(* IEC 61131-3 sources: daoli-st-library/DL_Device, 362 files *)

(* ---- FB_DL_AnalogInputRedundancySel.st ---- *)
(*==============================================================================
 * 组件名称 (Component)  : FB_DL_AnalogInputRedundancySel
 * 所属子库 (Sublibrary) : DL_Device
 * 当前版本 (Version)    : 1.0.0
 * 兼容性   (Platform)   : CODESYS 3.5 / TwinCAT 3 / 汇川 InoProShop / 施耐德 Machine Expert
 *                         仅依赖 IEC 61131-3 标准库（ABS / MAX / MIN），零厂商方言
 * 功能描述 (Function)   : 双路模拟量冗余选择（无扰切换 + 偏差监控 + 坏值剔除）：
 *                         ① 两路均有效且 |A − B| ≤ fDevTol → 输出两路均值，选通码 3；
 *                         ② 两路均有效但偏差超限 → **按上一拍选定通道保持**（无扰切换），
 *                            置 bDevAlarm 与信息码，绝不两侧来回跳；
 *                         ③ 仅一路有效（另一路非有限 / 超量程）→ 剔除坏路、使用好路，
 *                            bChanAValid / bChanBValid 回执逐路披露；
 *                         ④ **双路皆坏 → eFault**：输出保持**上一有效值**，bValid=FALSE，
 *                            故障级码配对置 bError，恢复路径唯一：bReset 且至少一路恢复有效。
 * 接口     (Interface)  : 输入 8 项（使能 / 复位 / 两路原值 / 偏差容差 / 量程上下限），
 *                         输出 10 项（输出值 / 选通码 / 偏差告警 / 两路有效回执 /
 *                         状态回执 / 有效性与故障码）。
 * 边界     (Boundary)   : ① 量程判定用 [fRangeMin, fRangeMax] 闭区间，超界即该路无效
 *                            （不做单侧饱和，饱和会把坏值伪装成合法满量程）；
 *                         ② 偏差容差以 1E-9 为下限钳位，防零容差导致恒告警；
 *                         ③ 双路皆坏时输出保持 fLastValid（上一有效值），若从未有过
 *                            有效值则输出 0 哨兵并披露（bValid=FALSE）；
 *                         ④ 非有限双判：NaN 用 x <> x，Inf 用 |x − x| > EPS 双侧直比；
 *                         ⑤ 零全局耦合（无 GVL / VAR_EXTERNAL / %I / %Q）。
 * 码表     (Codes)      : 本件占用 16#0004_1020 ~ 16#0004_102F 区间，实际使用 5 个：
 *                         1020 信息级 容差/量程参数钳位；1021 信息级 仅单路有效已剔除坏路；
 *                         1022 信息级 双路偏差超限已保持上一通道；1023 故障级 双路皆坏；
 *                         1024 故障级 非法状态兜底。信息级码永不置 bError。
 * 分工声明 (Scope)      : 与 FB_DL_AnalogTransmitter 分工：那件做单路原始量→工程量的
 *                         标定与滤波；本件只做「两路冗余仲裁与坏值剔除」，不做标定。
 * 开源溯源 (Origin)     : 开源溯源：原创实现（无外部代码引入）
 * 红线自检 (Redline)    : R1 ✓ 零 GVL / VAR_EXTERNAL ｜ R2 ✓ 零 %I/%Q/%M
 *                         R3 ✓ 纯 IEC 61131-3 ｜ R4 ✓ 非有限双判 + 容差钳位 + 无除零
 *                         R5 ✓ 声明逐行同行双语注释 ｜ R6 ✓ 五态 ENUM + CASE + ELSE
 *                         R7 ✓ 无定时器/边沿实例（N/A），无跨周期定时依赖
 * 修订历史 (Revision)   : 2026-11-23  v1.0.0  R77 首版
 * 验收向量 (Acceptance) :
 *   V1 两路 A=10.0、B=10.4、fDevTol=1.0：fOut=10.2、iSelChan=3、bDevAlarm=FALSE、bValid=TRUE。
 *   V2 承接 V1，随后 A=10.0、B=15.0（偏差 5.0 > 1.0）：fOut 保持通道 A 的 10.0、
 *      iSelChan=1、bDevAlarm=TRUE、uErrorId=16#0004_1022、bError=FALSE（信息级）。
 *   V3 A=NaN、B=12.0：bChanAValid=FALSE、bChanBValid=TRUE、fOut=12.0、iSelChan=2、
 *      uErrorId=16#0004_1021、bError=FALSE。
 *   V4 A=NaN、B 超量程（B=200.0，量程上限 100.0）：双路皆坏 → eStateOut=eFault、
 *      fOut 保持上一有效值、bValid=FALSE、uErrorId=16#0004_1023、bError=TRUE。
 *   V5 承接 V4，bReset 单拍且 A 恢复为 10.0：eStateOut 回 eAvg/eHoldA，bError=FALSE。
 *============================================================================*)

(*-----------------------------------------------------------------------------
 * 调用示例 (Instance guide)：
 *   声明于调用方 FB 的 VAR 区：fbRed : FB_DL_AnalogInputRedundancySel;
 *   每周期无条件调用：fbRed(bEnable := TRUE, bReset := xReset,
 *                           fChanA := stAi.fCh1, fChanB := stAi.fCh2,
 *                           fDevTol := 0.5, fRangeMin := 0.0, fRangeMax := 100.0);
 *   取用出口：fPv := fbRed.fOut;  IF NOT fbRed.bValid THEN 保持工艺安全动作。
 *   注意：iSelChan 为「上一拍选定通道」的唯一载体，请勿在外部改写。
 *----------------------------------------------------------------------------*)

(*-----------------------------------------------------------------------------
 * 枚举: E_DL_ArsState（归属 DL_Device，与 FB_DL_AnalogInputRedundancySel 同文件）
 * 含义: 冗余选择状态机的离散状态。eAvg 为双路均值相，eHoldA / eHoldB 为单路保持相，
 *       eFault 为双路皆坏的故障相（输出保持上一有效值）。
 *----------------------------------------------------------------------------*)
TYPE E_DL_ArsState :
(
    eInit  := 0,    // 首扫态：输出直接取可用路，建立首个有效值 / First scan: output takes a valid channel to build the first valid value
    eAvg   := 10,   // 均值态：两路有效且偏差合格，输出均值 / Averaging state: both valid and deviation within tolerance
    eHoldA := 20,   // 保持 A 态：仅 A 有效或偏差超限且上一拍选 A / Hold channel A, valid alone or deviation exceeded with A previously selected
    eHoldB := 30,   // 保持 B 态：仅 B 有效或偏差超限且上一拍选 B / Hold channel B, valid alone or deviation exceeded with B previously selected
    eFault := 99    // 故障相：双路皆坏，输出保持上一有效值，bValid=FALSE / Fault: both channels bad, holds last valid value
);
END_TYPE

(*==============================================================================
 * 功能块: FB_DL_AnalogInputRedundancySel
 * 调用约定: 每周期无条件调用一次；无定时器/边沿实例（R7 N/A），全部判据单拍完成。
 * 无扰语义: 通道间切换只发生在「上一拍选定通道仍然有效」的前提下；一旦选定通道
 *           失效才切到另一路，切回条件为原通道恢复有效（而非偏差合格），避免抖动。
 *============================================================================*)
FUNCTION_BLOCK FB_DL_AnalogInputRedundancySel
VAR_INPUT
    bEnable    : BOOL := FALSE;         // 使能，FALSE 时输出冻结并置 bValid=FALSE / Enable, FALSE freezes the output and clears bValid
    bReset     : BOOL := FALSE;         // 复位（电平有效），解除双路皆坏锁存 / Reset (level), clears the both-bad latch
    fChanA     : REAL := 0.0;           // A 路原始采样值 [EU] / Raw sample of channel A [EU]
    fChanB     : REAL := 0.0;           // B 路原始采样值 [EU] / Raw sample of channel B [EU]
    fDevTol    : REAL := 0.5;           // 两路允许偏差容差 [EU] / Allowed deviation between the two channels [EU]
    fRangeMin  : REAL := 0.0;           // 量程下限（闭区间）[EU] / Range lower bound, closed interval [EU]
    fRangeMax  : REAL := 100.0;         // 量程上限（闭区间）[EU] / Range upper bound, closed interval [EU]
END_VAR
VAR_OUTPUT
    fOut       : REAL;                  // 仲裁输出值（双路皆坏时保持上一有效值）[EU] / Arbitrated output, holds last valid on both-bad
    iSelChan   : INT;                   // 选通码：0=无 1=A 2=B 3=均值 [-] / Selection code: 0=none 1=A 2=B 3=mean
    bDevAlarm  : BOOL;                  // 双路偏差超限告警（信息级，不置 bError）/ Deviation alarm, info level, keeps bError FALSE
    bChanAValid: BOOL;                  // A 路有效回执（有限且在量程内）/ Channel A validity feedback, finite and in range
    bChanBValid: BOOL;                  // B 路有效回执（有限且在量程内）/ Channel B validity feedback, finite and in range
    eStateOut  : E_DL_ArsState;         // 状态机当前状态回执 [-] / Current state feedback
    bValid     : BOOL;                  // 输出可信标志，故障相为 FALSE / Output trustworthy flag, FALSE in the fault state
    bError     : BOOL;                  // 故障级标志，与 uErrorId 严格联动 / Fault-level flag, strictly coupled with uErrorId
    uErrorId   : UDINT;                 // 错误码，0 = 无码 / Error code, 0 = no code
END_VAR
VAR
    eState     : E_DL_ArsState;         // 内部状态 [-] / Internal state
    fDev       : REAL;                  // 两路实时偏差绝对值 [EU] / Absolute deviation between the two channels [EU]
    fLastValid : REAL;                  // 上一有效输出值，故障相保持用 [EU] / Last valid output, held in the fault state
    bHaveLast  : BOOL;                  // 是否已建立过有效值 / A valid value has been established
    bBothValid : BOOL;                  // 两路均有效 / Both channels valid
    bOnlyA     : BOOL;                  // 仅 A 有效 / Only channel A valid
    bOnlyB     : BOOL;                  // 仅 B 有效 / Only channel B valid
    bNoneValid : BOOL;                  // 两路皆无效 / Neither channel valid
    bDevOk     : BOOL;                  // 偏差在容差内 / Deviation inside tolerance
    bChanANaN  : BOOL;                  // A 路自反判 NaN 命中 / Channel A NaN by self-comparison
    bChanAInf  : BOOL;                  // A 路差自减判 Inf 命中 / Channel A infinity by self-subtraction
    bChanBNaN  : BOOL;                  // B 路自反判 NaN 命中 / Channel B NaN by self-comparison
    bChanBInf  : BOOL;                  // B 路差自减判 Inf 命中 / Channel B infinity by self-subtraction
    bFaultLatch: BOOL;                  // 双路皆坏锁存位 / Both-bad latch
    bRangeBad  : BOOL;                  // 量程参数非法标志 / Range parameter invalid flag
    fDevTolEff : REAL;                  // 钳位后的偏差容差 [EU] / Clamped deviation tolerance [EU]
    fRangeLo   : REAL;                  // 生效量程下限 [EU] / Effective range lower bound [EU]
    fRangeHi   : REAL;                  // 生效量程上限 [EU] / Effective range upper bound [EU]
    uInfoCode  : UDINT;                 // 信息级码暂存 / Info-level code scratch
END_VAR
VAR CONSTANT
    DL_ARS_OK    : UDINT := 16#0000_0000;  // 无码哨兵 / No-code sentinel
    DL_ARS_TOL   : REAL := 1.0E-9;         // 容差硬下限，防零容差恒告警 [EU] / Tolerance floor preventing permanent alarm [EU]
    DL_ARS_EPS   : REAL := 1.0E-9;         // 浮点比较容差（统一口径）/ Unified floating point comparison tolerance
    DL_ARS_ZERO  : REAL := 0.0;            // 零基准哨兵 / Zero reference sentinel
    DL_ARS_HALF  : REAL := 0.5;            // 均值折半系数 / Averaging half factor
    DL_ARS_RANGE_DEF : REAL := 100.0;      // 量程非法时的兜底上限 [EU] / Fallback upper bound when the range is invalid [EU]
END_VAR

(*------------------------------------------------------------------------------
 * 段 0｜参数域闸（不中断扫描）：量程必须 fRangeMax > fRangeMin，容差 ≥ 1E-9
 *      Parameter domain gate: range must be increasing, tolerance floored
 *-----------------------------------------------------------------------------*)
uInfoCode  := DL_ARS_OK;                                    // 信息码预置无码 / Preset no info code
bRangeBad  := FALSE;                                        // 量程非法标志预置 / Preset range-invalid flag FALSE

fDevTolEff := MAX(fDevTol, DL_ARS_TOL);                     // 容差下限钳位 [EU] / Tolerance floor [EU]
fRangeLo   := fRangeMin;                                    // 生效量程下限 [EU] / Effective lower bound [EU]
IF fRangeMax > fRangeMin THEN
    fRangeHi := fRangeMax;                                  // 量程合法原值生效 [EU] / Legal upper bound applied [EU]
ELSE
    fRangeHi   := fRangeLo + DL_ARS_RANGE_DEF;              // 量程倒挂：改用兜底上限，拒绝零宽量程 / Inverted range, fallback width
    bRangeBad  := TRUE;                                     // 记录量程非法 / Record the invalid range
    uInfoCode  := 16#0004_1020;                             // 信息级：量程参数已钳位 / Info: range parameter clamped
END_IF

(*------------------------------------------------------------------------------
 * 段 1｜逐路有效性判定：非有限（NaN 自反 / Inf 差自减）与超量程（闭区间）双闸
 *      Per-channel validity: non-finite double test plus closed-interval range gate
 *-----------------------------------------------------------------------------*)
bChanANaN := (fChanA <> fChanA);                                                          // A 路自反判 NaN / Channel A NaN by self-comparison
bChanAInf := ABS(fChanA - fChanA) > DL_ARS_EPS;                                           // A 路差自减判 Inf（双侧直比）/ Channel A infinity by self-subtraction
bChanAValid := NOT (bChanANaN OR bChanAInf)
               AND (fChanA >= fRangeLo) AND (fChanA <= fRangeHi);                          // A 路有效回执 / Channel A validity

bChanBNaN := (fChanB <> fChanB);                                                          // B 路自反判 NaN / Channel B NaN by self-comparison
bChanBInf := ABS(fChanB - fChanB) > DL_ARS_EPS;                                           // B 路差自减判 Inf（双侧直比）/ Channel B infinity by self-subtraction
bChanBValid := NOT (bChanBNaN OR bChanBInf)
               AND (fChanB >= fRangeLo) AND (fChanB <= fRangeHi);                          // B 路有效回执 / Channel B validity

bBothValid := bChanAValid AND bChanBValid;                  // 两路均有效 / Both valid
bOnlyA     := bChanAValid AND (NOT bChanBValid);            // 仅 A 有效 / Only A valid
bOnlyB     := bChanBValid AND (NOT bChanAValid);            // 仅 B 有效 / Only B valid
bNoneValid := (NOT bChanAValid) AND (NOT bChanBValid);      // 两路皆无效 / Neither valid

(* 偏差只在两路都有效时才有意义；任一路坏时偏差保持上一拍值（不拿坏值重算）*)
(* The deviation is meaningful only when both channels are valid, otherwise it is held *)
IF bBothValid THEN
    fDev := ABS(fChanA - fChanB);                           // 两路偏差绝对值 [EU] / Absolute deviation [EU]
END_IF
bDevOk := bBothValid AND (fDev <= fDevTolEff);             // 偏差合格判据 [EU] / Deviation predicate [EU]

(*------------------------------------------------------------------------------
 * 段 2｜双路皆坏锁存：置位在 eFault 判断处，解除路径唯一：bReset 且至少一路有效
 *      Both-bad latch: cleared only by reset with at least one channel valid again
 *-----------------------------------------------------------------------------*)
IF bFaultLatch THEN
    IF bReset AND (bChanAValid OR bChanBValid) THEN
        bFaultLatch := FALSE;                               // 唯一解除路径：复位且至少一路恢复有效 / Sole clear path
    END_IF
ELSIF bNoneValid AND bEnable THEN
    bFaultLatch := TRUE;                                    // 双路皆坏：锁存 / Both channels bad, latch it
END_IF

(*------------------------------------------------------------------------------
 * 段 3｜主状态机（红线 R6）：ENUM + CASE + ELSE 兜底
 *      Main state machine with enum, case coverage and ELSE interception
 *      出口预置：本件所有分支都显式给 fOut / iSelChan / bValid，无隐式保持
 *-----------------------------------------------------------------------------*)
CASE eState OF

    eInit:
        (* 首扫：不做仲裁，直接取可用路建立首个有效值 *)
        (* First scan: no arbitration, take an available channel to build the first valid value *)
        bDevAlarm := FALSE;                                 // 告警复位 / Alarm reset
        IF bBothValid THEN
            fOut       := (fChanA + fChanB) * DL_ARS_HALF;  // 两路可用取均值 [EU] / Both usable, take the mean [EU]
            iSelChan   := 3;                                // 选通码 3 = 均值 / Selection code three, mean
            fLastValid := fOut;                             // 建立首个有效值 / Build the first valid value
            bHaveLast  := TRUE;                             // 有效值已建立 / Valid value established
            bValid     := TRUE;                             // 输出可信 / Output trustworthy
            eState     := eAvg;                             // 进均值相 / Enter the averaging state
        ELSIF bOnlyA THEN
            fOut       := fChanA;                           // 仅 A 可用 [EU] / Only A usable [EU]
            iSelChan   := 1;                                // 选通码 1 = A / Selection code one, A
            fLastValid := fOut;                             // 建立首个有效值 / Build the first valid value
            bHaveLast  := TRUE;                             // 有效值已建立 / Valid value established
            bValid     := TRUE;                             // 输出可信 / Output trustworthy
            eState     := eHoldA;                           // 进保持 A 相 / Enter hold A
        ELSIF bOnlyB THEN
            fOut       := fChanB;                           // 仅 B 可用 [EU] / Only B usable [EU]
            iSelChan   := 2;                                // 选通码 2 = B / Selection code two, B
            fLastValid := fOut;                             // 建立首个有效值 / Build the first valid value
            bHaveLast  := TRUE;                             // 有效值已建立 / Valid value established
            bValid     := TRUE;                             // 输出可信 / Output trustworthy
            eState     := eHoldB;                           // 进保持 B 相 / Enter hold B
        ELSIF bEnable THEN
            fOut      := fLastValid;                        // 双路皆坏：保持上一有效值（可能仍是 0 哨兵）/ Both bad, hold the last valid value
            iSelChan  := 0;                                 // 无选定通道 / No selected channel
            bValid    := FALSE;                             // 输出不可信 / Output untrustworthy
            bDevAlarm := FALSE;                             // 偏差判据不可得，不置告警 / Deviation unavailable, no alarm
            eState    := eFault;                            // 进故障相 / Enter the fault state
        ELSE
            fOut      := fLastValid;                        // 未使能：输出冻结 / Not enabled, output frozen
            iSelChan  := 0;                                 // 无选定通道 / No selected channel
            bValid    := FALSE;                             // 输出不可信 / Output untrustworthy
        END_IF

    eAvg:
        (* 均值相：两路仍有效且偏差合格才保持；偏差超限则保持上一拍选定通道 *)
        (* Averaging state: keep averaging while the deviation is fine, else hold the previous channel *)
        IF bNoneValid THEN
            fOut      := fLastValid;                        // 双路皆坏：保持上一有效值 / Both bad, hold the last valid value
            iSelChan  := 0;                                 // 无选定通道 / No selected channel
            bValid    := FALSE;                             // 输出不可信 / Output untrustworthy
            bDevAlarm := FALSE;                             // 偏差判据不可得 / Deviation unavailable
            eState    := eFault;                            // 进故障相 / Enter the fault state
        ELSIF bOnlyA THEN
            fOut       := fChanA;                           // 剔除坏路 B，用 A [EU] / Drop B, use A [EU]
            iSelChan   := 1;                                // 选通码 1 = A / Selection code one, A
            fLastValid := fOut;                             // 刷新上一有效值 / Refresh the last valid value
            bHaveLast  := TRUE;                             // 有效值已建立 / Valid value established
            bValid     := TRUE;                             // 输出可信 / Output trustworthy
            bDevAlarm  := FALSE;                            // 单路运行不属偏差告警 / Single-channel run is not a deviation alarm
            uInfoCode  := 16#0004_1021;                     // 信息级：仅单路有效已剔除坏路 / Info: single channel valid, bad one dropped
            eState     := eHoldA;                           // 进保持 A 相 / Enter hold A
        ELSIF bOnlyB THEN
            fOut       := fChanB;                           // 剔除坏路 A，用 B [EU] / Drop A, use B [EU]
            iSelChan   := 2;                                // 选通码 2 = B / Selection code two, B
            fLastValid := fOut;                             // 刷新上一有效值 / Refresh the last valid value
            bHaveLast  := TRUE;                             // 有效值已建立 / Valid value established
            bValid     := TRUE;                             // 输出可信 / Output trustworthy
            bDevAlarm  := FALSE;                            // 单路运行不属偏差告警 / Single-channel run is not a deviation alarm
            uInfoCode  := 16#0004_1021;                     // 信息级：仅单路有效已剔除坏路 / Info: single channel valid, bad one dropped
            eState     := eHoldB;                           // 进保持 B 相 / Enter hold B
        ELSIF bDevOk THEN
            fOut       := (fChanA + fChanB) * DL_ARS_HALF;  // 偏差合格：取均值 [EU] / Deviation fine, take the mean [EU]
            iSelChan   := 3;                                // 选通码 3 = 均值 / Selection code three, mean
            fLastValid := fOut;                             // 刷新上一有效值 / Refresh the last valid value
            bHaveLast  := TRUE;                             // 有效值已建立 / Valid value established
            bValid     := TRUE;                             // 输出可信 / Output trustworthy
            bDevAlarm  := FALSE;                            // 告警复位 / Alarm reset
        ELSE
            (* 偏差超限：无扰保持上一拍选定通道；均值相无历史通道时按 A 保持（口径写死）*)
            (* Deviation exceeded: hold the previous channel; from the mean state default to A *)
            fOut       := fChanA;                           // 保持 A 通道值（均值相缺历史时的固定口径）[EU] / Hold A, fixed policy from the mean state [EU]
            iSelChan   := 1;                                // 选通码 1 = A / Selection code one, A
            fLastValid := fOut;                             // 刷新上一有效值 / Refresh the last valid value
            bHaveLast  := TRUE;                             // 有效值已建立 / Valid value established
            bValid     := TRUE;                             // 输出可信 / Output trustworthy
            bDevAlarm  := TRUE;                             // 偏差超限告警置位 / Deviation alarm set
            uInfoCode  := 16#0004_1022;                     // 信息级：偏差超限已保持上一通道 / Info: deviation exceeded, previous channel held
            eState     := eHoldA;                           // 进保持 A 相 / Enter hold A
        END_IF

    eHoldA:
        (* 保持 A 相：A 仍有效即继续；A 失效则切 B；两路皆坏进故障相 *)
        (* Hold A: continue while A is valid, switch to B when A fails, fault when both bad *)
        IF bNoneValid THEN
            fOut      := fLastValid;                        // 双路皆坏：保持上一有效值 / Both bad, hold the last valid value
            iSelChan  := 0;                                 // 无选定通道 / No selected channel
            bValid    := FALSE;                             // 输出不可信 / Output untrustworthy
            bDevAlarm := FALSE;                             // 偏差判据不可得 / Deviation unavailable
            eState    := eFault;                            // 进故障相 / Enter the fault state
        ELSIF bChanAValid THEN
            fOut       := fChanA;                           // 保持 A 路 [EU] / Hold channel A [EU]
            iSelChan   := 1;                                // 选通码 1 = A / Selection code one, A
            fLastValid := fOut;                             // 刷新上一有效值 / Refresh the last valid value
            bHaveLast  := TRUE;                             // 有效值已建立 / Valid value established
            bValid     := TRUE;                             // 输出可信 / Output trustworthy
            IF bBothValid AND (NOT bDevOk) THEN
                bDevAlarm := TRUE;                          // 两路都在但偏差超限：维持告警 / Both valid but deviating, keep the alarm
                uInfoCode := 16#0004_1022;                  // 信息级：偏差超限保持通道 / Info: deviation exceeded, channel held
            ELSE
                bDevAlarm := FALSE;                         // 偏差回落清除告警 / Alarm cleared when the deviation settles
            END_IF
        ELSE
            fOut       := fChanB;                           // A 失效切 B（B 此时必然有效）[EU] / A failed, switch to B, which must be valid [EU]
            iSelChan   := 2;                                // 选通码 2 = B / Selection code two, B
            fLastValid := fOut;                             // 刷新上一有效值 / Refresh the last valid value
            bHaveLast  := TRUE;                             // 有效值已建立 / Valid value established
            bValid     := TRUE;                             // 输出可信 / Output trustworthy
            bDevAlarm  := FALSE;                            // 单路运行不属偏差告警 / Single-channel run is not a deviation alarm
            uInfoCode  := 16#0004_1021;                     // 信息级：仅单路有效已剔除坏路 / Info: single channel valid, bad one dropped
            eState     := eHoldB;                           // 进保持 B 相 / Enter hold B
        END_IF

    eHoldB:
        (* 保持 B 相：B 仍有效即继续；B 失效则切 A；两路皆坏进故障相 *)
        (* Hold B: continue while B is valid, switch to A when B fails, fault when both bad *)
        IF bNoneValid THEN
            fOut      := fLastValid;                        // 双路皆坏：保持上一有效值 / Both bad, hold the last valid value
            iSelChan  := 0;                                 // 无选定通道 / No selected channel
            bValid    := FALSE;                             // 输出不可信 / Output untrustworthy
            bDevAlarm := FALSE;                             // 偏差判据不可得 / Deviation unavailable
            eState    := eFault;                            // 进故障相 / Enter the fault state
        ELSIF bChanBValid THEN
            fOut       := fChanB;                           // 保持 B 路 [EU] / Hold channel B [EU]
            iSelChan   := 2;                                // 选通码 2 = B / Selection code two, B
            fLastValid := fOut;                             // 刷新上一有效值 / Refresh the last valid value
            bHaveLast  := TRUE;                             // 有效值已建立 / Valid value established
            bValid     := TRUE;                             // 输出可信 / Output trustworthy
            IF bBothValid AND (NOT bDevOk) THEN
                bDevAlarm := TRUE;                          // 两路都在但偏差超限：维持告警 / Both valid but deviating, keep the alarm
                uInfoCode := 16#0004_1022;                  // 信息级：偏差超限保持通道 / Info: deviation exceeded, channel held
            ELSE
                bDevAlarm := FALSE;                         // 偏差回落清除告警 / Alarm cleared when the deviation settles
            END_IF
        ELSE
            fOut       := fChanA;                           // B 失效切 A（A 此时必然有效）[EU] / B failed, switch to A, which must be valid [EU]
            iSelChan   := 1;                                // 选通码 1 = A / Selection code one, A
            fLastValid := fOut;                             // 刷新上一有效值 / Refresh the last valid value
            bHaveLast  := TRUE;                             // 有效值已建立 / Valid value established
            bValid     := TRUE;                             // 输出可信 / Output trustworthy
            bDevAlarm  := FALSE;                            // 单路运行不属偏差告警 / Single-channel run is not a deviation alarm
            uInfoCode  := 16#0004_1021;                     // 信息级：仅单路有效已剔除坏路 / Info: single channel valid, bad one dropped
            eState     := eHoldA;                           // 进保持 A 相 / Enter hold A
        END_IF

    eFault:
        (* 故障相：输出保持上一有效值，bValid=FALSE；恢复路径唯一：bReset 且至少一路有效 *)
        (* Fault: hold the last valid value, recover only via reset with one valid channel *)
        fOut      := fLastValid;                            // 保持上一有效值（从未有过则为 0 哨兵）/ Hold the last valid value
        iSelChan  := 0;                                     // 无选定通道 / No selected channel
        bValid    := FALSE;                                 // 输出不可信 / Output untrustworthy
        bDevAlarm := FALSE;                                 // 偏差判据不可得，不置告警 / Deviation unavailable, no alarm
        IF (NOT bEnable) THEN
            eState := eInit;                                // 失能回首扫态 / Disable returns to init
        ELSIF (NOT bFaultLatch) AND bChanAValid THEN
            eState := eHoldA;                               // 复位后 A 恢复有效 / A recovered after reset
        ELSIF (NOT bFaultLatch) AND bChanBValid THEN
            eState := eHoldB;                               // 复位后 B 恢复有效 / B recovered after reset
        END_IF

    ELSE
        (* 非法状态拦截：任何未定义枚举值一律进故障相并置兜底码 *)
        (* Illegal state interception: undefined enum values go to fault with a fallback code *)
        eState    := eFault;                                // 强制回故障相 / Force back to the fault state
        fOut      := fLastValid;                            // 输出保持上一有效值 / Output holds the last valid value
        iSelChan  := 0;                                     // 无选定通道 / No selected channel
        bValid    := FALSE;                                 // 输出不可信 / Output untrustworthy
        bDevAlarm := FALSE;                                 // 不置偏差告警 / No deviation alarm
        uInfoCode := 16#0004_1024;                          // 故障级：非法状态兜底 / Fault: illegal state fallback

END_CASE

(*------------------------------------------------------------------------------
 * 段 4｜无扰冻结：未使能时输出冻结在上一有效值（不跟随输入）
 *      Bumpless freeze: while disabled the output stays on the last valid value
 *-----------------------------------------------------------------------------*)
IF NOT bEnable THEN
    IF bHaveLast THEN
        fOut := fLastValid;                                 // 冻结在上一有效值 / Freeze on the last valid value
    ELSE
        fOut := DL_ARS_ZERO;                                // 从未有过有效值：输出 0 哨兵 / Never valid, emit the zero sentinel
    END_IF
    bValid    := FALSE;                                     // 冻结相输出不可信 / Frozen output is not trustworthy
    bDevAlarm := FALSE;                                     // 冻结相不产生告警 / No alarm while frozen
END_IF

(*------------------------------------------------------------------------------
 * 段 5｜故障码统一出口（故障级锁存回放，信息级不置 bError）
 *      Unified code outlet: fault codes replayed latched, info codes never raise bError
 *-----------------------------------------------------------------------------*)
IF bFaultLatch THEN
    uErrorId := 16#0004_1023;                               // 故障级：双路皆坏 / Fault: both channels bad
    bError   := TRUE;                                       // 故障级码配对置位 / Paired fault flag set
ELSIF uInfoCode = 16#0004_1024 THEN
    uErrorId := 16#0004_1024;                               // 故障级：非法状态兜底 / Fault: illegal state fallback
    bError   := TRUE;                                       // 故障级码配对置位 / Paired fault flag set
ELSE
    uErrorId := uInfoCode;                                  // 信息级码或 0 / Info code or zero
    bError   := FALSE;                                      // 信息级不置故障标志 / Info level never raises the fault flag
END_IF

eStateOut := eState;                                        // 状态回执单一出口 / State feedback through a single outlet
END_FUNCTION_BLOCK

(* ---- FB_DL_AnalogSignalHealth.st ---- *)
// ==============================================================================
// 组件名 Component  : FB_DL_AnalogSignalHealth
// 分类   Category   : DL_Device
// 前缀   Naming     : FB_DL_ ｜ b/f/e/t/u 类型前缀制（R265）
// 版本   Version    : 1.0.0
// 复杂度 Complexity  : 中
// 功能   Purpose    : 4-20mA 模拟量信号健康诊断：断线（< 3.6 mA）、超上限
//                      （> fSatHigh）、低限（fSatLow ≤ 值 < 3.6 之外的
//                      低带口径见边界三）、卡滞（变化率绝对值持续
//                      <= fStuckBand 超 tStuck）；报警锁存至 bReset 上升沿，
//                      沿脉冲单拍。供变送器回路质量监视与预测性维护。
// 开源溯源 Origin    : 西门子 LGF 分类语义借鉴，clean-room 重写（LGF
//                      Process Diagnostics「模拟量断线 / 饱和监视」分类学
//                      口径借鉴，只借骨不抄肉，判据与实现零代码复制）
// 许可证 License    : MIT
// 参考   Reference  : IEC 61131-3:2013 §6.6 TON / R_TRIG 语义；NAMUR
//                      NE43 信号电平分级公开条款（借 3.6/4/20/20.5 mA
//                      分级语义，不抄文）
// 平台   Platform   : 纯 IEC 61131-3（TON / R_TRIG / LREAL 比较），三平台通用
// 依赖   Depends    : 仅 Standard.library（TON / R_TRIG 属标准件）
// 分工声明 Split     : FB_DL_SignalStuckWatch（通用卡滞监视）/ FB_DL_Analog
//                      Transmitter（模拟量变换）与本件互引；本件为 4-20mA
//                      回路专属健康分级（NE43 口径 + 回路卡滞三合一），
//                      通用信号冻结监视归 SignalStuckWatch（R216）。
// 归属 Ownership     : E_DL_AshHealth 属主为本文件（全库唯一定义，R264）；
//                      引用件只引用不重声明。
// ------------------------------------------------------------------
// 边界 Boundary     :
//   一 TON 无条件刷新（R7）：tonStuck 于段 0 顶层调用，IN 串「有变化即
//      重置」口径——IN := 变化率绝对值 <= fStuckBand（有变化时 IN 为
//      FALSE 计时自清，卡滞即「无变化持续超窗」）；首拍 / 复位后
//      _bPrevValid = FALSE 不计时（防假前值参与变化率）；
//   二 判据分级（R190 归因唯一，独立码位）：fMa 非有限 → eInvalid
//      （bValid = FALSE 通道，无码位）；fMa < 3.6 → eWireBreak（断线）；
//      fMa >= 3.6 且 fMa < fSatLow → eSatLow（低限）；fMa > fSatHigh →
//      eSatHigh（超上限）；其余正常带内 tonStuck.Q → eStuck（卡滞）；
//      以上皆否 → eOk；
//   三 低限口径声明：3.6 mA 硬断线阈值与 fSatLow 组态阈值分离——
//      fSatLow 默认 3.6（与硬阈值重合），调用方可上调 fSatLow 收紧
//      低带；fSatLow 下调低于 3.6 时低限带被硬阈值吸收（合法组态）；
//   四 报警锁存：_bAlarmLatch 置位后保持至 bReset 上升沿（锁存解除式
//      可达自证：输入引脚恒可达，R152）；首报码 _uErrLatch 锁存回放
//      （FB33-1：不在故障态按当下输入重新推断）；bAlarmEdge 单拍
//      （新报警沿，已锁存期不再发）；
//   五 组态守卫（防御性补码，R272 逐项点名）：fSatLow >= fSatHigh、
//      fSatLow / fSatHigh / fStuckBand 非有限、fStuckBand < 0、
//      tStuck <= 0 任一成立 → eHealth = eInvalid、bValid = FALSE、
//      报警锁存（故障级 0735）；
//   六 卡滞窗与报警锁存互锁：_bAlarmLatch 期间 tonStuck.IN 强制 FALSE
//      （复位沿同拍不重锁，FB50-1），复位后 _bPrevValid 清零重练；
//   七 失能（bEn = FALSE）语义写死（R303 离相清零）：eHealth 回 eOk、
//      报警锁存 / 码锁存清零、bValid = FALSE（失能不是故障）；
//   八 无除法；无全局、无外部变量、无物理地址；无状态机 CASE
//      （IF 判据链，末位 ELSE 兜底为 eOk）。
// 错误码 Codes      :
//   16#0003_0201【信息级】断线（fMa < 3.6 mA，NE43 口径）→ eWireBreak
//   16#0003_0202【信息级】超上限（fMa > fSatHigh）→ eSatHigh
//   16#0003_0203【信息级】低限（3.6 ≤ fMa < fSatLow）→ eSatLow
//   16#0003_0204【信息级】卡滞（变化率 <= fStuckBand 持续 tStuck）→ eStuck
//   16#0003_0735【故障级】组态非法（fSatLow >= fSatHigh / 参数非有限 /
//                fStuckBand < 0 / tStuck <= 0）→ eInvalid + bValid = FALSE
//   注：0201~0204 段位按本轮任务定稿启用（信息级，经 eErr / bAlarm
//   通道表达）；fMa 非有限走 eInvalid 无码位（bValid = FALSE 通道）。
//   0201~0204 四码分立依据（R90）：处置人不同（断线查接线、超限查
//   量程组态、低限查供电、卡滞查管路 / 变送器膜片），场景互斥可还原。
// 验收 Acceptance   :
//   算法已证（脚本）：未跑 ｜ 编译器已证（三平台）：未跑
//   V1 fMa = 3.0 → eWireBreak + 码 0201 + bAlarm 锁存
//   V2 fMa = 21.0 → eSatHigh + 码 0202；fMa = 3.7（fSatLow = 4.0）→ eSatLow
//   V3 fMa 恒 12.000 ± 0.01 超 10s → eStuck + 码 0204
//   V4 fMa 恒定但 < 3.6 → 断线优先（卡滞窗被门控不计时）
//   V5 fMa = NaN → eInvalid + bValid = FALSE（无码位）
//   V6 bReset 上升沿 → 锁存清零、卡滞计时重练（_bPrevValid 清零）
//   V7 bEn = FALSE → 全出口清零回 eOk（R303）
//   V8 fSatLow = 25（>= fSatHigh）→ 0735 + eInvalid
// 修订记录 Revision  :
//   2026-11-22  v1.0.0  R65 首版（批 3 · 序号 9，LGF Process Diagnostics 补口）
// ==============================================================================
TYPE E_DL_AshHealth :
(
    eOk        := 0,  // 健康带内 / ok, the signal in the healthy band
    eWireBreak := 10, // 断线：fMa < 3.6 mA（NE43 口径）/ the wire break under the hard threshold
    eSatHigh   := 20, // 超上限：fMa > fSatHigh / the saturation above the configured high
    eSatLow    := 30, // 低限：3.6 <= fMa < fSatLow / the low limit under the configured low
    eStuck     := 40, // 卡滞：变化率持续不超带超窗 / the stuck value through the window
    eInvalid   := 50  // 无效：输入非有限或组态非法 / invalid, a non finite input or configuration
);
END_TYPE

FUNCTION_BLOCK FB_DL_AnalogSignalHealth
VAR_INPUT
    fMa        : LREAL;         // 实测电流 [mA]（4-20mA 回路）/ the measured current in milliamps
    bEn        : BOOL := TRUE;  // 使能 [-]，FALSE 时出口清零回 eOk（R303）/ the enable
    fSatLow    : LREAL := 3.6;  // 低限阈值 [mA]，须 < fSatHigh / the low limit threshold
    fSatHigh   : LREAL := 20.5; // 超上限阈值 [mA]，NE43 口径默认 20.5 / the saturation high threshold
    fStuckBand : LREAL := 0.05; // 卡滞变化带 [mA]，变化率绝对值 <= 此值视为无变化 / the stuck band of the rate
    tStuck     : TIME := T#10S; // 卡滞判定窗 [毫秒]，须 > 0 / the stuck window, above zero
    bReset     : BOOL := FALSE; // 报警复位电平，上升沿清锁存（边界四解除式）/ the reset level, its rising edge releases the latch
END_VAR
VAR_OUTPUT
    eHealth    : E_DL_AshHealth := E_DL_AshHealth.eOk; // 健康状态出口 [状态] / the health outlet
    bAlarm     : BOOL := FALSE; // 报警锁存 [-]，任一非 eOk 状态置位至复位 / the latched alarm
    bAlarmEdge : BOOL := FALSE; // 新报警沿脉冲 [-]，单拍有效 / the new alarm edge pulse, single scan
    bValid     : BOOL := FALSE; // 判据可用 [-]，输入非有限或组态非法为 FALSE / the criteria usable flag
    eErr       : UDINT := 16#0000_0000; // 错误码，0 = 正常（首报码锁存回放）/ the error code, zero is ok
END_VAR
VAR
    _fPrevMa     : LREAL := 0.0;  // 前拍 mA 快照 [mA]（卡滞变化率基准）/ the previous scan snapshot of fMa
    _bPrevValid  : BOOL := FALSE; // 前值有效标志 [-]（首拍 / 复位后不参与变化率）/ the previous value valid flag
    _bAlarmLatch : BOOL := FALSE; // 报警锁存副本 [-]（仅复位沿清除）/ the alarm latch copy
    _uErrLatch   : UDINT := 16#0000_0000; // 首报码锁存 [码]（复位沿清除，FB33-1）/ the latched first report code
    _bAlarmNew   : BOOL := FALSE; // 本拍新报警标志 [-]（沿脉冲源，单拍）/ the new alarm flag of this scan
    _eHealthInt  : E_DL_AshHealth := E_DL_AshHealth.eOk; // 健康状态内部判定 [状态] / the internal health verdict
    _uCodeNow    : UDINT := 16#0000_0000; // 本拍判据码 [码] / the verdict code of this scan
    _bMaBad      : BOOL;          // fMa 非有限标志（逐拍重算）/ the input fault flag
    _bCfgBad     : BOOL;          // 组态非法标志（逐拍重算）/ the configuration fault flag
    _bInBand     : BOOL;          // 处于正常工作带 [-]（卡滞计时前提）/ the in band flag, the stuck timer premise
    _bDeltaSmall : BOOL;          // 变化率不超带 [-]（卡滞计时条件）/ the small rate flag
    rtReset      : R_TRIG;        // 复位沿实例，段 0 无条件刷新（R7）/ the reset edge instance refreshed unconditionally
    tonStuck     : TON;           // 卡滞窗定时器，段 0 无条件刷新 / the stuck window timer refreshed unconditionally
END_VAR
VAR CONSTANT
    DL_ASH_WIRE  : LREAL := 3.6;            // 硬断线阈值 [mA]（NE43 口径）/ the hard wire break threshold
    DL_ASH_FMAX  : LREAL := 1.0E30;         // 非有限筛查幅值上限 [mA] / the finiteness screening cap
    DL_ASH_TIME0 : TIME := T#0S;            // 时间零常量 [毫秒] / the time zero constant
    DL_ASH_ZEROU : UDINT := 16#0000_0000;   // 码零常量 / the code zero constant
    DL_ASH_E_WIRE  : UDINT := 16#0003_0201; // 信息级：断线 / the wire break code
    DL_ASH_E_SATHI : UDINT := 16#0003_0202; // 信息级：超上限 / the saturation high code
    DL_ASH_E_SATLO : UDINT := 16#0003_0203; // 信息级：低限 / the low limit code
    DL_ASH_E_STUCK : UDINT := 16#0003_0204; // 信息级：卡滞 / the stuck code
    DL_ASH_E_CFG   : UDINT := 16#0003_0735; // 故障级：组态非法 / the configuration fault code
END_VAR

// 段 0｜定时器与沿实例无条件周期刷新（禁入分支，R7）/ segment 0, the unconditional refresh
rtReset(CLK := bReset);          // 复位沿 / the reset edge
_bMaBad := (fMa <> fMa) OR ((fMa - fMa) <> 0.0) OR (ABS(fMa) > DL_ASH_FMAX); // 输入非有限（NaN 自反判 + Inf 差值自反判 + 幅值上界，R272）/ the input non finite
_bCfgBad := (fSatLow >= fSatHigh)                                        // 低限不低于上限 / the low limit above the high
         OR (fSatLow <> fSatLow) OR ((fSatLow - fSatLow) <> 0.0) OR (ABS(fSatLow) > DL_ASH_FMAX)     // fSatLow 非有限 / fSatLow non finite
         OR (fSatHigh <> fSatHigh) OR ((fSatHigh - fSatHigh) <> 0.0) OR (ABS(fSatHigh) > DL_ASH_FMAX) // fSatHigh 非有限 / fSatHigh non finite
         OR (fStuckBand < 0.0)                                           // 变化带为负 / a negative band
         OR (fStuckBand <> fStuckBand) OR ((fStuckBand - fStuckBand) <> 0.0) OR (ABS(fStuckBand) > DL_ASH_FMAX) // fStuckBand 非有限 / fStuckBand non finite
         OR (tStuck <= DL_ASH_TIME0);                                    // 卡滞窗非正 / a non positive window
_bInBand := (NOT _bMaBad) AND (NOT _bCfgBad) AND (fMa >= DL_ASH_WIRE) AND (fMa >= fSatLow) AND (fMa <= fSatHigh); // 正常工作带（卡滞计时前提，边界二）/ the healthy band, the stuck timer premise
_bDeltaSmall := _bPrevValid AND (ABS(fMa - _fPrevMa) <= fStuckBand); // 变化率不超带（有变化时为 FALSE 计时自清，边界一）/ the rate within the band
tonStuck(IN := bEn AND _bInBand AND (NOT _bAlarmLatch) AND _bDeltaSmall, PT := tStuck); // 卡滞窗计时（串使能 / 带 / 锁存门控，FB50-1；锁存期 IN 强制 FALSE 防复位同拍重锁，边界六）/ the stuck window with the full gating

// 段 1｜单拍量预清零 + 复位沿作用域（R256 / R311）/ segment 1, the preset and the reset edge scope
bAlarmEdge := FALSE;             // 沿脉冲预清零（单拍信息位）/ preset the edge pulse false
IF rtReset.Q THEN                // 复位沿（作用域声明：清双锁存 + 重练卡滞计时，R311）/ the reset edge with the declared scope
    _bAlarmLatch := FALSE;       // 清报警锁存（唯一解除路径，边界四自证可达）/ clear the alarm latch
    _uErrLatch := DL_ASH_ZEROU;  // 清首报码锁存 / clear the latched code
    _bPrevValid := FALSE;        // 前值失效（卡滞计时重练，防旧基线误判）/ invalidate the previous value
    _fPrevMa := 0.0;             // 前值显式清零 [mA] / clear the previous value explicitly
END_IF

// 段 2｜失能分支：出口清零回 eOk，不 faults（R303 离相清零声明行）/ segment 2, the disabled branch
IF NOT bEn THEN                  // 失能 / disabled
    _eHealthInt := E_DL_AshHealth.eOk; // 强制健康态 / force the healthy state
    _bAlarmLatch := FALSE;       // 清报警锁存（使能断开 ≠ 信号故障）/ clear the alarm latch
    _uErrLatch := DL_ASH_ZEROU;  // 清码锁存 / clear the latched code
    _bPrevValid := FALSE;        // 前值失效（重新使能后重练）/ invalidate the previous value
    eHealth := _eHealthInt;      // 状态出口 / the health outlet
    bAlarm := FALSE;             // 报警位复位 / the alarm bit resets
    bAlarmEdge := FALSE;         // 沿脉冲复位 / the edge pulse resets
    bValid := FALSE;             // 失能即不可用 / not usable while disabled
    eErr := DL_ASH_ZEROU;        // 失能不发码 / no code while disabled
    RETURN;                      // 早退 / early return
END_IF

// 段 3｜判据分级链（边界二 / 五：R190 归因唯一，末位 ELSE 兜底 eOk）/ segment 3, the verdict chain
IF _bCfgBad THEN                 // 组态非法优先（故障级 0735）/ the configuration fault first
    _eHealthInt := E_DL_AshHealth.eInvalid; // 无效态 / the invalid state
    _uCodeNow := DL_ASH_E_CFG;   // 故障级码 / the fault code
ELSIF _bMaBad THEN               // 输入非有限 / a non finite input
    _eHealthInt := E_DL_AshHealth.eInvalid; // 无效态 / the invalid state
    _uCodeNow := DL_ASH_ZEROU;   // 无码位（bValid = FALSE 通道表达，边界二）/ no code, the validity channel speaks
ELSIF fMa < DL_ASH_WIRE THEN     // 硬断线阈值之下（NE43 口径）/ under the hard wire break threshold
    _eHealthInt := E_DL_AshHealth.eWireBreak; // 断线态 / the wire break state
    _uCodeNow := DL_ASH_E_WIRE;  // 信息级 0201 / the wire break code
ELSIF fMa < fSatLow THEN         // 低限带（fMa >= 3.6 已由上分支证明）/ the low limit band
    _eHealthInt := E_DL_AshHealth.eSatLow;   // 低限态 / the low limit state
    _uCodeNow := DL_ASH_E_SATLO; // 信息级 0203 / the low limit code
ELSIF fMa > fSatHigh THEN        // 超上限 / over the high threshold
    _eHealthInt := E_DL_AshHealth.eSatHigh;  // 超上限态 / the saturation state
    _uCodeNow := DL_ASH_E_SATHI; // 信息级 0202 / the saturation code
ELSIF tonStuck.Q THEN            // 卡滞超窗（正常带内才有资格判，边界二 / 六）/ stuck through the window
    _eHealthInt := E_DL_AshHealth.eStuck;    // 卡滞态 / the stuck state
    _uCodeNow := DL_ASH_E_STUCK; // 信息级 0204 / the stuck code
ELSE                             // 兜底：健康 / the fallback, healthy
    _eHealthInt := E_DL_AshHealth.eOk;       // 健康态 / the healthy state
    _uCodeNow := DL_ASH_ZEROU;   // 无码 / no code
END_IF

// 段 4｜报警锁存与首报码（边界四：锁存回放，FB33-1）/ segment 4, the alarm latch and the first report code
_bAlarmNew := FALSE;             // 新报警标志预清零 / preset the new alarm flag false
IF _eHealthInt <> E_DL_AshHealth.eOk THEN // 判据非健康 / the verdict not healthy
    IF NOT _bAlarmLatch THEN     // 首次报警 / a first alarm
        _bAlarmNew := TRUE;      // 置新报警标志（沿脉冲源，单拍）/ raise the new alarm flag
        _uErrLatch := _uCodeNow; // 首报码锁存（此后回放，不按当下输入重推断）/ latch the first code for the replay
    END_IF
    _bAlarmLatch := TRUE;        // 报警锁存至复位沿 / latch the alarm to the reset edge
END_IF

// 段 5｜统一出口（名实双出口同源，R191）/ segment 5, the unified outlet
eHealth := _eHealthInt;          // 状态出口 / the health outlet
bAlarm := _bAlarmLatch;          // 报警位与锁存同源 / the alarm bit from the latch
bAlarmEdge := _bAlarmNew;        // 沿脉冲单拍（已锁存期不再发）/ the single scan edge pulse
bValid := (NOT _bMaBad) AND (NOT _bCfgBad); // 判据可用（无输入 / 组态故障）/ usable without faults
IF _bAlarmLatch THEN             // 报警锁存回放优先 / the latched code replays first
    eErr := _uErrLatch;          // 首报码回放 / replay the latched code
ELSE                             // 无报警 / no alarm
    eErr := DL_ASH_ZEROU;        // 正常 / ok
END_IF

// 段 6｜前拍快照更新（边界一：仅有限值更新，非有限保旧值）/ segment 6, the previous value update
IF NOT _bMaBad THEN              // 输入有限才更新基准 / update the baseline only on a finite input
    _fPrevMa := fMa;             // 前拍快照刷新 [mA] / refresh the snapshot
    _bPrevValid := TRUE;         // 前值有效 / the previous value valid
END_IF
END_FUNCTION_BLOCK

(* ---- FB_DL_AxiolineDiagLatch.st ---- *)
(*==============================================================================
 * 组件名称 (Component)  : FB_DL_AxiolineDiagLatch
 * 所属子库 (Sublibrary) : DL_Device
 * 当前版本 (Version)    : 1.0.1
 * 组件分类 (Category)   : 功能块（FUNCTION_BLOCK）· 设备诊断 · 总线位域解析
 * 兼容性   (Platform)   : CODESYS 3.5 / TwinCAT 3 / 汇川 InoProShop / Schneider
 *                         Machine Expert；仅位与运算与标准 TON / R_TRIG
 * 功能描述 (Function)   : 把本地总线的诊断状态寄存器位域与诊断参数寄存器
 *                         （错误码加槽号）解析为工程师可直接读的分级诊断：
 *                         总线级、模块级、通道级三档，加首出故障槽号、错误码、
 *                         防抖事件计数与锁存和复位语义。
 * 位序声明 (Bit layout) : 本块常量位序为自有定义：PF 为 bit0、PW 为 bit1、
 *                         BUS 为 bit2、RUN 为 bit3、ACT 为 bit4、RDY 为 bit5、
 *                         SYSFAIL 为 bit6。现场寄存器的高低字节拼接由调用方在
 *                         IO 映射层完成，本块不做任何字节序猜测（跨平台歧义禁令），
 *                         头注释即为对照表，接线变更只改 IO 层。
 * 槽号特例 (Slot cases) : 槽号 0 表示无位置信息，输出 -1；槽号 128 表示
 *                         「无法定位」，原值保留供 HMI 直接显示定位失败，
 *                         绝不折算成 128 号槽；大于 127 且不等于 128 属非法，
 *                         按无位置处理并置信息级码。
 * 首出锁存 (First-out)  : 首个稳定成立的诊断被锁存后，后续新诊断不覆盖首出，
 *                         这正是排故需要的因果顺序；确认（Ack）只清显示位，
 *                         不清锁存；只有复位（Reset）才清锁存。此语义与
 *                          FB_DL_InterlockMatrix 的首出思想同源但独立实现。
 * 设计要点 (Key notes)  : ① 分级判定先判致命：系统故障或（总线错误且总线未
 *                           就绪）优先于一切外围故障，避免 HMI 只看到一条
 *                           「模块故障」而漏掉真正的总线掉站；
 *                         ② 防抖：只有状态稳定超过稳定窗才计入事件，瞬断不会
 *                           让事件计数暴涨，也不会误锁首出；
 *                         ③ 未使能时清实时诊断位但保留锁存历史：检修断电前
 *                           仍能在 HMI 上看到最后一个首出槽号，不丢现场证据；
 *                         ④ 事件计数只增不减，复位不清（计数值是台账），
 *                           只清锁存与首出。
 * 开源溯源 (Origin)     : plcnext-community。参考 PLCnext 官方在线帮助公开的
 *                         本地总线诊断系统变量语义（外围故障、外围警告、总线
 *                         错误、运行、组态就绪、总线就绪、系统故障七个位义，
 *                         诊断参数寄存器给错误码、扩展参数给错误位置槽号，
 *                         无法定位用 128 表示）。只借位语义与「错误码加槽号」
 *                         参数域，寄存器字宽、位序、枚举、码位与状态机 100%
 *                         自有，输入一律经引脚注入，不绑定任何厂商系统变量，
 *                         clean-room，不构成衍生作品。
 * 依赖     (Depends)    : 无 DL_ 内部依赖；仅 Standard.library 的 TON / R_TRIG
 * 故障码表 (Error codes):
 *   16#0003_013B【信息级】槽号非法（大于 127 且不等于 128），按无位置处理
 *   16#0003_013C【信息级】诊断块未使能，实时位已清零、锁存保留
 *   16#0003_02F4【故障级】诊断位有效但错误码为 0（状态与参数寄存器不自洽）
 *   16#0003_02F5【故障级】非法状态兜底
 *   16#0003_02F6【故障级】总线就绪丢失超时（诊断有效而模块就绪长时间为假）
 * 验收向量 (Acceptance) :
 *   V1 状态字 16#0001（外围故障）/ 错误码 16#0102 / 槽号 3 → 稳定 200 毫秒后
 *      等级为故障、首出槽号 3、首出码 16#0102、事件计数 1
 *   V2 随后再来槽号 7 错误码 16#0204 → 首出槽号仍为 3（首因不覆盖）
 *   V3 槽号 128 → 首出槽号 128（不得变成 -1）
 *   V4 状态字 16#0044（总线错误加系统故障）→ 等级为致命，而非故障
 *   V5 状态字 100 毫秒内抖动 5 次 → 事件计数只加 1
 *   V6 复位一拍 → 首出槽号 -1、事件计数保持、事件码清零
 * 红线自检 (Redline)    : R1 零全局变量表与外部变量引用 ｜ R2 零物理地址直写
 *                         R3 纯 IEC 61131-3 ｜ R4 位运算无越界、无除法、无浮点
 *                         R5 全变量中英双语同行注释 ｜ R6 ENUM 加 CASE 加 ELSE 兜底
 *                         R7 TON 与两个 R_TRIG 全部在 CASE 之外无条件刷新
 * 修订历史 (Revision)   :
 *   2026-11-15  v1.0.0  首版入库（Round 10 · T1-7 PLCnext 开组）
 *   2026-11-15  v1.0.1  R10 终审修复三处：
 *                       R-FIX-1【严重】确认屏蔽计数在同一拍内先装载后递减，
 *                       屏蔽长度恒为 0，bAckDiag 完全无效（规格要求确认沿清
 *                       显示位）；改为装载拍不递减，确认当拍起生效；
 *                       R-FIX-2【中等】未使能时 eMonitor 仍可锁存并累加事件，
 *                       与「未使能只清实时位、保留历史」矛盾；锁存条件加使能；
 *                       R-FIX-3【注释级】事件台账段落原文把 uEventCnt 描述为
 *                       「故障发生了几次」，与「锁存后不覆盖、复位前不再加一」
 *                       的实际行为不符，已按实际语义改写（R12 向量/描述自洽）。
 *============================================================================*)

(*------------------------------------------------------------------------------
 * 枚举: E_DL_DiagLevel（诊断等级，归属本功能块并同文件发布）
 *-----------------------------------------------------------------------------*)
TYPE E_DL_DiagLevel :
(
    eNone  := 0,     // 无诊断：全部诊断位为零 / No diagnostic, every bit clear
    eWarn  := 10,    // 警告：外围警告位有效，可继续生产 / Warning, production may continue
    eFault := 20,    // 故障：外围故障位有效，模块或通道级硬件问题 / Fault, module or channel level hardware issue
    eFatal := 30     // 致命：系统故障或总线掉站，须立即停机排故 / Fatal, system failure or bus loss, stop the machine
);
END_TYPE

(*------------------------------------------------------------------------------
 * 枚举: E_DL_DiagFsm（本块状态机，归属本功能块并同文件发布）
 *-----------------------------------------------------------------------------*)
TYPE E_DL_DiagFsm :
(
    eIdle    := 0,   // 待机：未使能或尚未建立监视 / Idle, disabled or not monitoring yet
    eMonitor := 10,  // 监视中：实时解析诊断，未锁存 / Monitoring, live diagnostics parsed, nothing latched
    eLatched := 20,  // 已锁存首出：新诊断不覆盖 / Latched, subsequent diagnostics do not overwrite
    eFault   := 99   // 故障：状态与参数不自洽或非法状态 / Fault, inconsistency or illegal state
);
END_TYPE

(*==============================================================================
 * 逐拍推演 (Cycle-by-cycle trace)：
 *   场景 A 单个外围故障（状态字 16#0001，错误码 16#0102，槽号 3）
 *     拍 1 位域解析出外围故障，原始聚合为真，槽号解析为 3
 *          稳定窗重新计时，稳定标志仍假，不锁存，等级为故障
 *     中途每拍状态字与错误码不变，稳定窗持续计时
 *     稳定窗到（约 200 毫秒后，取决于任务周期）
 *          稳定标志为真且等级非无，未锁存过，锁存槽号 3 与码 16#0102，
 *          事件计数加 1，转已锁存态；错误码非零，不置 02F4
 *   场景 B 首出不覆盖（随后槽号 7，错误码 16#0204）
 *     已锁存态下新诊断只被观测，不覆盖已锁存槽号与码，首出仍为 3
 *   场景 C 无法定位（槽号 128）
 *     解析结果保持 128（不折算成 128 号槽，也不变成无位置），供 HMI 直接
 *     显示「定位失败」
 *   场景 D 致命优先（状态字 16#0044，即总线错误加系统故障，模块未就绪）
 *     分级先判致命条件，等级取致命，不再落到故障档
 *   场景 E 抖动 5 次（100 毫秒内状态字反复变化）
 *     稳定窗每次被重置，始终未到，事件计数一次都不加；待状态稳定后才加 1
 *   场景 F 复位一拍
 *     锁存清除、槽号回负一、码清零；事件计数保持（台账不清）
 *============================================================================*)

(*==============================================================================
 * 位序对照表 (Bit order cross reference)：
 *   位号   本库常量名        含义              现场常见语义        判读建议
 *   bit0   DL_BIT_PF        外围故障          模块或通道硬件错    先看槽号
 *   bit1   DL_BIT_PW        外围警告          非致命，可继续生产  记录趋势
 *   bit2   DL_BIT_BUS       总线错误          总线通信异常        结合就绪位
 *   bit3   DL_BIT_RUN       数据传输中        数据正在交换        正常运行应为真
 *   bit4   DL_BIT_ACT       组态就绪          组态已生效          启动前应为真
 *   bit5   DL_BIT_RDY       总线就绪          总线可用            启动前应为真
 *   bit6   DL_BIT_SYSFAIL   系统故障          设备级致命故障      立即停机
 *   说明：本表是调用方在 IO 层拼字节时的唯一依据；若现场寄存器的高低位与
 *   本表相反，请在 IO 层做字节交换后再送进本块，不要改本块的常量。
 *============================================================================*)

(*==============================================================================
 * 事件台账语义 (Event ledger)：
 *   uEventCnt 是累计锁存次数，只在「本轮锁存成立」那一拍加一：同一故障持续
 *   存在期间不会每拍累加，锁存之后到复位之前到来的新诊断也不会再加——即它
 *   计数的是「已锁存的首出事件轮次」，不是每一类故障各自的发生次数。需要
 *   逐类次数统计时，请在上层按 uFirstCode 分类后自行累加，不要改本块的
 *   加一条件（改了会让「首因不覆盖」这条排故原则失效）。
 *   uFirstCode 与 uFirstSlot 记录的是本轮锁存中最早捕获的那一条，后续
 *   新故障不会覆盖它们，这与「首出优先」的电气排故原则一致：先解释
 *   第一个故障，后面的往往是它的连锁反应。
 *============================================================================*)

FUNCTION_BLOCK FB_DL_AxiolineDiagLatch
VAR_INPUT
    bEnable      : BOOL := TRUE;     // 使能，FALSE 时清实时诊断位但保留锁存 [-] / Enable, FALSE clears live bits but keeps the latch
    uStatusWord  : WORD;             // 诊断状态寄存器位域，字节拼接由 IO 层完成 [位串] / Diagnostic status register, byte order merged by the IO layer
    uErrCode     : WORD;             // 诊断参数寄存器：错误码 [代码] / Diagnostic parameter register, the error code
    uErrSlot     : USINT;            // 扩展参数寄存器：错误位置槽号，0 与 128 为特例 [槽] / Error location slot, zero and 128 are special
    bModuleReady : BOOL;             // 总线就绪反馈，等价总线就绪位，冗余校验用 [-] / Bus ready feedback, redundant with the ready bit
    bAckDiag     : BOOL;             // 诊断确认，上升沿清显示位但不清锁存 [-] / Diagnostic acknowledge, clears display bits only
    bReset       : BOOL;             // 复位锁存与首出，上升沿有效 [-] / Reset the latch and the first-out record
END_VAR
VAR_OUTPUT
    bBusError    : BOOL;             // 总线级故障（总线错误位）[-] / Bus level fault
    bPeriphFault : BOOL;             // 外围故障（外围故障位），模块或通道硬件错 [-] / Peripheral fault
    bPeriphWarn  : BOOL;             // 外围警告（外围警告位）[-] / Peripheral warning
    bSysFail     : BOOL;             // 系统故障（系统故障位）[-] / System failure
    bDiagActive  : BOOL;             // 任一诊断有效，聚合位供 HMI 单点使用 [-] / Any diagnostic active, an aggregate bit for the HMI
    eLevel       : E_DL_DiagLevel;   // 诊断等级（无 / 警告 / 故障 / 致命）[-] / Diagnostic level
    nFirstSlot   : INT := -1;        // 首出故障槽号，-1 表示无，128 表示无法定位 [槽] / First-out slot, -1 none, 128 unlocatable
    uFirstCode   : WORD;             // 首出故障错误码，与槽号同拍锁存 [代码] / First-out error code latched together with the slot
    nEventCnt    : UDINT;            // 诊断事件累计次数，去抖后计数，复位不清 [次] / Debounced event counter, never cleared by reset
    bLatchFull   : BOOL;             // 锁存已满（首出保持，需复位）[-] / Latch occupied, needs a reset
    uErrorId     : UDINT;            // 事件码，0 = 无事件 / Event code, 0 = no event
END_VAR
VAR
    fbTrigAck    : R_TRIG;           // 确认沿检测，CASE 之外无条件刷新 [-] / Rising edge detector for the acknowledge input
    fbTrigReset  : R_TRIG;           // 复位沿检测，CASE 之外无条件刷新 [-] / Rising edge detector for the reset input
    fbDebounce   : TON;              // 诊断稳定窗计时，CASE 之外无条件刷新 [-] / Diagnostic stabilisation timer
    bInit        : BOOL := FALSE;    // 首扫标志，初值 FALSE，判据 NOT bInit（R19 范式）[-] / First-scan flag
    bLatched     : BOOL;             // 首出锁存有效 [-] / TRUE when the first-out record is latched
    nSlotLatch   : INT := -1;        // 锁存槽号 [槽] / Latched slot number
    uCodeLatch   : WORD;             // 锁存错误码 [代码] / Latched error code
    eState       : E_DL_DiagFsm := E_DL_DiagFsm.eIdle;  // 状态机 / State machine
    uPrevStatus  : WORD;             // 上拍状态字，用于变化检测 [位串] / Previous status word for change detection
    bDebIn       : BOOL;             // 稳定窗输入条件，先算后调以免条件调用实例 [-] / Stabilisation input condition computed before the call
    bRawActive   : BOOL;             // 原始诊断位聚合（未去抖）[-] / Raw aggregate of the diagnostic bits before debouncing
    bStable      : BOOL;             // 去抖后的稳定诊断标志 [-] / Debounced diagnostic flag
    nSlotParsed  : INT;              // 槽号解析结果 [槽] / Parsed slot number
    eLevelRaw    : E_DL_DiagLevel;   // 未去抖的原始等级 [-] / Raw diagnostic level before debouncing
    nAckMute     : INT;              // 确认屏蔽计数，确认后抑制显示若干拍 [拍] / Acknowledge mute counter
END_VAR
VAR CONSTANT
    DL_BIT_PF      : WORD := 16#0001;    // 外围故障位（本库自有位序，bit0）[位串] / Peripheral fault bit
    DL_BIT_PW      : WORD := 16#0002;    // 外围警告位（bit1）[位串] / Peripheral warning bit
    DL_BIT_BUS     : WORD := 16#0004;    // 总线错误位（bit2）[位串] / Bus error bit
    DL_BIT_RUN     : WORD := 16#0008;    // 数据传输中位（bit3）[位串] / Data transfer running bit
    DL_BIT_ACT     : WORD := 16#0010;    // 组态就绪位（bit4）[位串] / Configuration active bit
    DL_BIT_RDY     : WORD := 16#0020;    // 总线就绪位（bit5）[位串] / Bus ready bit
    DL_BIT_SYSFAIL : WORD := 16#0040;    // 系统故障位（bit6）[位串] / System failure bit
    DL_SLOT_UNLOC  : USINT := 128;       // 无法定位标志 [槽] / Unlocatable marker
    DL_SLOT_NONE   : USINT := 0;         // 无位置信息 [槽] / No location information
    DL_SLOT_MAX    : INT := 127;         // 有效槽号上限 [槽] / Highest valid slot number
    DL_DEB_TIME    : TIME := T#200MS;    // 诊断稳定窗 [毫秒] / Diagnostic stabilisation window
    DL_ACK_MUTE    : INT := 1;           // 确认后抑制显示的拍数 [拍] / Cycles to mute the display after an acknowledge
END_VAR

(*------------------------------------------------------------------------------
 * 段 1｜沿检测无条件刷新（R7 红线）
 *      Edge detection refreshed unconditionally
 *-----------------------------------------------------------------------------*)
fbTrigAck(CLK := bAckDiag);
fbTrigReset(CLK := bReset);

(*------------------------------------------------------------------------------
 * 段 2｜首扫初始化（R19 唯一合法范式）
 *      First-scan initialisation with the canonical R19 pattern
 *-----------------------------------------------------------------------------*)
IF NOT bInit THEN
    bLatched    := FALSE;
    nSlotLatch  := -1;
    uCodeLatch  := 16#0000;
    nEventCnt   := 0;
    uErrorId    := 16#0000_0000;
    eState      := E_DL_DiagFsm.eIdle;
    uPrevStatus := 16#0000;
    nAckMute    := 0;
    bInit       := TRUE;                 // 首扫只做一次
END_IF

(*------------------------------------------------------------------------------
 * 段 3｜位域解析：状态字按自有位序拆七个位，不做字节序猜测
 *      Bit field decode using the library-owned bit order, no byte order guessing
 *-----------------------------------------------------------------------------*)
IF (uStatusWord AND DL_BIT_PF) <> 16#0000 THEN
    bPeriphFault := TRUE;
ELSE
    bPeriphFault := FALSE;
END_IF

IF (uStatusWord AND DL_BIT_PW) <> 16#0000 THEN
    bPeriphWarn := TRUE;
ELSE
    bPeriphWarn := FALSE;
END_IF

IF (uStatusWord AND DL_BIT_BUS) <> 16#0000 THEN
    bBusError := TRUE;
ELSE
    bBusError := FALSE;
END_IF

IF (uStatusWord AND DL_BIT_SYSFAIL) <> 16#0000 THEN
    bSysFail := TRUE;
ELSE
    bSysFail := FALSE;
END_IF

IF bBusError OR bPeriphFault OR bPeriphWarn OR bSysFail THEN
    bRawActive := TRUE;
ELSE
    bRawActive := FALSE;
END_IF

(*------------------------------------------------------------------------------
 * 段 4｜槽号解析（三特例写死）
 *      Slot parsing with three hard-coded special cases
 *-----------------------------------------------------------------------------*)
IF uErrSlot = DL_SLOT_NONE THEN
    nSlotParsed := -1;                       // 无位置信息
ELSIF uErrSlot = DL_SLOT_UNLOC THEN
    nSlotParsed := 128;                      // 无法定位：原值保留，不伪装成槽号
ELSIF USINT_TO_INT(uErrSlot) <= DL_SLOT_MAX THEN
    nSlotParsed := USINT_TO_INT(uErrSlot);   // 1 到 127：有效槽号
ELSE
    nSlotParsed := -1;                       // 大于 127 且不等于 128：非法
    uErrorId    := 16#0003_013B;
END_IF

(*------------------------------------------------------------------------------
 * 段 5｜稳定窗计时（红线：定时器在 CASE 之外无条件刷新）
 *      Stabilisation timer refreshed unconditionally outside the CASE
 *      输入条件为「原始诊断有效」或「状态字发生变化」，任一成立即重新计时
 *-----------------------------------------------------------------------------*)
IF bRawActive OR (uStatusWord <> uPrevStatus) THEN
    bDebIn := TRUE;
ELSE
    bDebIn := FALSE;
END_IF
fbDebounce(IN := bDebIn, PT := DL_DEB_TIME);
bStable := fbDebounce.Q;

(*------------------------------------------------------------------------------
 * 段 6｜分级判定（先判致命，顺序不得调整）
 *      Level classification, fatal first, the order must not be changed
 *-----------------------------------------------------------------------------*)
IF bSysFail OR (bBusError AND (NOT bModuleReady)) THEN
    eLevelRaw := E_DL_DiagLevel.eFatal;
ELSIF bPeriphFault THEN
    eLevelRaw := E_DL_DiagLevel.eFault;
ELSIF bPeriphWarn THEN
    eLevelRaw := E_DL_DiagLevel.eWarn;
ELSE
    eLevelRaw := E_DL_DiagLevel.eNone;
END_IF

(*------------------------------------------------------------------------------
 * 段 7｜主状态机（ENUM 加 CASE，含 ELSE 兜底）
 *      Main state machine with an ELSE fallback branch
 *-----------------------------------------------------------------------------*)
CASE eState OF
    E_DL_DiagFsm.eIdle:
        IF bEnable THEN
            eState := E_DL_DiagFsm.eMonitor;
        END_IF

    E_DL_DiagFsm.eMonitor:
        (* 稳定成立的诊断才锁首出：瞬断不计事件，避免事件计数暴涨
           未使能时不得锁存新事件：使能失败/检修期间只保留历史，不污染台账 *)
        IF bEnable AND bStable AND (eLevelRaw <> E_DL_DiagLevel.eNone) THEN
            IF NOT bLatched THEN
                nSlotLatch := nSlotParsed;
                uCodeLatch := uErrCode;
                bLatched   := TRUE;
                nEventCnt  := nEventCnt + 1;
                eState     := E_DL_DiagFsm.eLatched;
                IF uErrCode = 16#0000 THEN
                    uErrorId := 16#0003_02F4;    // 状态位与参数寄存器不自洽
                END_IF
            END_IF
        END_IF

    E_DL_DiagFsm.eLatched:
        (* 首出锁定：新诊断不覆盖首出槽号与首出码，只保留因果顺序中的首因 *)
        IF NOT bEnable THEN
            eState := E_DL_DiagFsm.eIdle;
        END_IF

    E_DL_DiagFsm.eFault:
        (* 故障：仅复位沿可退，复位处理在段 8 中执行，此处保持故障码 *)
        uErrorId := 16#0003_02F5;

    ELSE
        eState   := E_DL_DiagFsm.eFault;
        uErrorId := 16#0003_02F5;
END_CASE

(*------------------------------------------------------------------------------
 * 段 8｜确认与复位（复位放在锁存之后，保证复位当拍首出即为 -1）
 *      Acknowledge and reset, reset placed after latching so it wins this cycle
 *-----------------------------------------------------------------------------*)
IF fbTrigAck.Q THEN
    nAckMute := DL_ACK_MUTE;             // 确认拍：装载屏蔽长度，当拍不清零
ELSIF nAckMute > 0 THEN
    nAckMute := nAckMute - 1;            // 非确认拍才递减，否则屏蔽长度恒为 0
END_IF

IF fbTrigReset.Q THEN
    bLatched   := FALSE;
    nSlotLatch := -1;
    uCodeLatch := 16#0000;
    uErrorId   := 16#0000_0000;
    IF bEnable THEN
        eState := E_DL_DiagFsm.eMonitor;
    ELSE
        eState := E_DL_DiagFsm.eIdle;
    END_IF
END_IF

(*------------------------------------------------------------------------------
 * 段 9｜总线就绪丢失超时（故障级）：诊断有效而模块就绪长时间为假
 *      Bus ready loss watchdog: diagnostics active while the module stays unready
 *      判定放在状态机之后，只置码不改状态，避免与首出锁存争夺状态迁移权
 *-----------------------------------------------------------------------------*)
IF bStable AND bRawActive AND (NOT bModuleReady) THEN
    uErrorId := 16#0003_02F6;
END_IF

(*------------------------------------------------------------------------------
 * 段 10｜输出每拍重写（R27）：未使能时清实时位、保留锁存历史
 *      Outputs rewritten every cycle; disabled clears live bits but keeps history
 *-----------------------------------------------------------------------------*)
IF bEnable THEN
    IF bRawActive AND (nAckMute = 0) THEN
        bDiagActive := TRUE;
    ELSE
        bDiagActive := FALSE;
    END_IF
    eLevel     := eLevelRaw;
    uFirstCode := uCodeLatch;            // 首出码与首出槽号同源，锁存后每拍重写
ELSE
    bBusError    := FALSE;
    bPeriphFault := FALSE;
    bPeriphWarn  := FALSE;
    bSysFail     := FALSE;
    bDiagActive  := FALSE;
    eLevel       := E_DL_DiagLevel.eNone;
    uFirstCode   := uCodeLatch;          // 锁存历史保留，便于未使能时排故
    uErrorId     := 16#0003_013C;        // 信息级：诊断块未使能
END_IF

nFirstSlot := nSlotLatch;                // 首出槽号每拍重写，复位后自然变 -1
bLatchFull := bLatched;
uPrevStatus := uStatusWord;              // 变化检测基准更新，必须在解析之后
END_FUNCTION_BLOCK

(* ---- FB_DL_CassetteBcdLabel.st ---- *)
(*==============================================================================
 * 组件名称 (Component)  : FB_DL_CassetteBcdLabel
 * 所属子库 (Sublibrary) : DL_Device
 * 当前版本 (Version)    : 1.0.0
 * 兼容性   (Platform)   : CODESYS 3.5+ / TwinCAT 3 / 汇川 InoProShop / 施耐德 Machine Expert
 *                         仅依赖 Standard.library（TON / R_TRIG / LEN），零厂商私有库
 * 功能描述 (Function)   : 花篮 BCD 拨码标签机联动。
 *                         把批次号（0..9999）编成 4 位 BCD 拨码，驱动标签机打印，再用扫码枪回读
 *                         校验"打出来的标签"与"拨码值"一致，形成闭环；不一致或打印超时即锁存。
 *                         三段语义：
 *                           ① **拨码生成**：数值 → 四位十进制 → 打包 BCD（移位量取常量 0/4/8/12，
 *                              恒小于 WORD 位宽 16），并做**逐位 BCD 校验**（每位 ≤ 9，由十进制拆分
 *                              结构性保证，另设反解校验以覆盖"外部写入 BCD 字"的通道）；
 *                           ② **扫码枪语义**：回读串逐字符转数字并校验字符合法（'0'..'9'），
 *                              非法字符即判 eScanFormat；
 *                           ③ **打印同步握手**：打印脉冲单拍 → 等 bPrintDone → 扫码校验 → 结果脉冲。
 *                         **忙时拒新任务**：打印窗口内收到新的生成请求只置 bBusyReject（信息级），
 *                         不打断当前任务（打断会产生半张标签，比排队更糟）。
 *                         验收向量：
 *                           ① 批次 1234 → uBcd = 16#1234，四位数字 4/3/2/1
 *                           ② 回读 "1234" → 校验通过，bLabelOk 单拍
 *                           ③ 回读 "12X4" → eScanFormat 锁存（非法字符）
 *                           ④ 回读 "1235" → eScanMismatch 锁存（数值不一致）
 *                           ⑤ 打印窗口内再次请求生成 → bBusyReject 单拍，当前任务不受影响
 * 接口     (Interface)  : 入 iLotNo 批次号（0..9999）、bGenReq 生成沿、bPrintDone 打印完成、
 *                         sScanCode 扫码回读串、bScanValid 回读有效、tPrintTo 打印超时、bReset 复位沿；
 *                         出 uBcdPacked 打包 BCD、abDigits 四位数字（1=个 … 4=千）、bPrintCmd 打印脉冲（单拍）、
 *                         bLabelOk 标签校验通过脉冲（单拍）、bBusy 打印中、bBusyReject 忙拒单拍、
 *                         bLabelFail 标签失败锁存、eState 相、eCause 成因、bError 故障标志。
 * 边界     (Boundary)   : ① **属主边界（写死）：本件只做"拨码编码 + 打印握手 + 扫码校验"，
 *                         不驱动打印头/拨码继电器、不解析标签条码的厂商前缀**（属设备驱动与协议件）；
 *                         ② **BCD 半字节校验**：位宽 16 恰 4 个半字节，校验域 k=0..3 完整覆盖，
 *                         头注释声明"不做越界半字节校验"（R57：越域半字节不存在而非非法）；
 *                         ③ **域闸**：iLotNo 越 0..9999 → 拒生成 + eLotBad（信息级）；
 *                         ④ **打印超时 TON**：tonPrint 段 0 无条件调用，IN 串 (NOT _bFault)，
 *                         故障期不累计，复位同拍不会立即重锁（R252）；
 *                         ⑤ **锁存解除式**：bLabelFail / eFault 仅由 bReset 上升沿解除（R228B），
 *                         bReset 为外部引脚、恒可达；
 *                         ⑥ 零全局耦合、零物理地址。
 * 分工声明 (Scope)      : 本件只管"花篮拨码标签联动"。不接管：IV 测试仪设定值导出
 *                         （属 FB_DL_IvBcdExport）、标签模板排版（属标签设计侧）、
 *                         花篮工艺履历（属追溯件）。
 * 来源标签 (Source Tag) : ROADMAP 空勾真缺口 P2（花篮 BCD 标签联动，自研 clean-room）
 * 码表     (Codes)      : 本件不占用任何全局数字码位（零码位范式 R297）；诊断由 BOOL + ENUM 出口承担。
 * 红线自检 (Redline)    : R1 ✓ 零 GVL/VAR_EXTERNAL ｜ R2 ✓ 零 %I/%Q/%M ｜ R3 ✓ 纯 IEC 61131-3
 *                         R4 ✓ 域闸 + 字符域校验 + 常量移位 + 超时 TON ｜ R5 ✓ 声明逐行同行双语注释
 *                         R6 ✓ ENUM+CASE 含 ELSE 兜底 ｜ R7 ✓ TON/三 R_TRIG 段 0 无条件刷新
 * 修订历史 (Revision)   : 2026-11-19  v1.0.0  R47 首版（批次 4 · 序号 18）
 *==============================================================================*)

TYPE E_DL_CblState :
(
    eIdle    := 0,    // 待机相（等生成请求） / Idle, awaiting a generation request
    ePrinting:= 10,   // 打印中（等打印完成） / Printing, awaiting completion
    eVerify  := 20,   // 校验相（等扫码回读） / Verifying, awaiting the scan read-back
    eFault   := 90    // 故障相（等复位） / Fault, awaiting reset
);
END_TYPE

TYPE E_DL_CblCause :
(
    eNone        := 0,   // 无异常 / No anomaly
    eLotBad      := 1,   // 批次号越域（信息级，拒生成） / Lot number out of range, info level
    eBusyReject  := 2,   // 忙时拒新任务（信息级） / Busy, new request rejected, info level
    ePrintTimeout:= 3,   // 打印超时（锁存） / Print timeout, latched
    eScanFormat  := 4,   // 回读含非法字符（锁存） / Illegal character in the read-back, latched
    eScanMismatch:= 5,   // 回读与拨码不一致（锁存） / Read-back mismatch, latched
    eCfgIllegal  := 6,   // 组态非法（超时非正） / Illegal configuration
    ePhaseBad    := 7    // 非法相位兜底 / Illegal phase fallback
);
END_TYPE

FUNCTION_BLOCK FB_DL_CassetteBcdLabel
VAR_INPUT
    iLotNo     : INT := 0;                 // 批次号，域 0..9999 [-] / Lot number, domain 0..9999
    bGenReq    : BOOL := FALSE;            // 生成请求沿 [-] / Generation request edge
    bPrintDone : BOOL := FALSE;            // 打印完成（当拍电平） [-] / Print finished, level
    sScanCode  : STRING[15] := '';         // 扫码回读串 [-] / Scan read-back string
    bScanValid : BOOL := FALSE;            // 回读有效（当拍电平） [-] / Read-back valid, level
    tPrintTo   : TIME := T#10S;            // 打印超时，域 > T#0S [ms] / Print timeout, > T#0S
    bReset     : BOOL := FALSE;            // 故障复位沿 [-] / Fault reset edge
END_VAR
VAR_OUTPUT
    uBcdPacked : WORD := 16#0000;                        // 打包 BCD 字 [BCD] / Packed BCD word
    abDigits   : ARRAY[1..4] OF BYTE;                    // 四位数字（1=个,2=十,3=百,4=千） [-] / Four digits
    bPrintCmd  : BOOL := FALSE;                          // 打印脉冲（单拍） [-] / Print pulse, single scan
    bLabelOk   : BOOL := FALSE;                          // 标签校验通过脉冲（单拍） [-] / Label verified pulse
    bBusy      : BOOL := FALSE;                          // 打印/校验中 [-] / Busy
    bBusyReject: BOOL := FALSE;                          // 忙拒单拍 [-] / Busy rejection, single scan
    bLabelFail : BOOL := FALSE;                          // 标签失败锁存（等复位） [-] / Label failure, latched
    eState     : E_DL_CblState := E_DL_CblState.eIdle;   // 相出口 [-] / Phase outlet
    eCause     : E_DL_CblCause := E_DL_CblCause.eNone;   // 成因出口（R190 归因唯一） [-] / Cause outlet
    bError     : BOOL := FALSE;                          // 故障标志（仅故障级成因） [-] / Error flag, fault level only
END_VAR
VAR
    _eState   : E_DL_CblState := E_DL_CblState.eIdle;    // 内部相（CASE 唯一写入目标） / Internal phase
    _eCause   : E_DL_CblCause := E_DL_CblCause.eNone;    // 成因锁存量 / Latched cause
    _bFault   : BOOL := FALSE;                           // 故障锁存位 / Latched fault bit
    _bFail    : BOOL := FALSE;                           // 标签失败锁存位 / Latched label-failure bit
    _uBcd     : WORD := 16#0000;                         // 打包工作值 [BCD] / Packing working value
    _iWork    : INT := 0;                                // 十进制拆分工作值 [-] / Decimal split working value
    _iVal     : INT := 0;                                // 回读串解析出的数值 [-] / Value parsed from the read-back
    _iPos     : INT := 0;                                // 回读串字符位置 / Character position in the read-back
    _iLen     : INT := 0;                                // 回读串长度 [字符] / Read-back length
    _iDigit   : INT := 0;                                // 当前字符代表的数字值（0..9） [-] / Digit value of the current character
    sChr      : STRING[1] := '';                         // 当前单字符（用于 '0'..'9' 判等） [-] / Current single character
    _bPrintCmd: BOOL := FALSE;                           // 打印脉冲内部位（单拍） / Internal print pulse
    _bLabelOk : BOOL := FALSE;                           // 校验通过内部位（单拍） / Internal verified pulse
    _bBusyRej : BOOL := FALSE;                           // 忙拒内部位（单拍） / Internal busy-rejection flag
    _bFmtBad  : BOOL := FALSE;                           // 回读格式结论 [-] / Read-back format result
    _bCfgBad  : BOOL := FALSE;                           // 组态非法当拍量 / Illegal configuration this scan
    tonPrint  : TON;                                     // 打印超时实例，段 0 无条件调用 / Print timeout instance
    rtGen     : R_TRIG;                                  // 生成沿实例，段 0 无条件调用 / Generation edge instance
    rtReset   : R_TRIG;                                  // 复位沿实例，段 0 无条件调用 / Reset edge instance
END_VAR
VAR CONSTANT
    DL_CBL_LOT_MAX : INT := 9999;        // 批次号上限（四位十进制） [-] / Lot upper bound
    DL_CBL_SH4     : INT := 4;           // 十位左移量（恒 < 16，R48） [bit] / Tens shift
    DL_CBL_SH8     : INT := 8;           // 百位左移量（恒 < 16，R48） [bit] / Hundreds shift
    DL_CBL_SH12    : INT := 12;          // 千位左移量（恒 < 16，R48） [bit] / Thousands shift
    DL_CBL_MSK     : WORD := 16#000F;    // 半字节掩码（非事件码，头注释声明） [bit] / Nibble mask, not an event code
    DL_CBL_CHR_MAX : INT := 15;          // 回读串长度硬上限（与 STRING[15] 同源） [字符] / Hard length ceiling
END_VAR

(* —— 段 0：组态闸 + TON 与两沿无条件周期刷新（R228A；IN 串故障否决，R252） —— *)
_bCfgBad := (tPrintTo <= T#0S);                                             // 打印超时须为正 / Timeout must be positive
rtGen(CLK := bGenReq);                                                      // 生成沿 / Generation edge
rtReset(CLK := bReset);                                                     // 复位沿 / Reset edge
tonPrint(IN := (_eState = E_DL_CblState.ePrinting) AND (NOT _bFault), PT := tPrintTo);   // 打印超时 / Print timeout

(* —— 段 1：单拍量预清零（锁存量 _eCause/_bFault/_bFail 不入清单，R107） —— *)
_bPrintCmd := FALSE;                                                        // 打印脉冲预清 / Print pulse preset
_bLabelOk  := FALSE;                                                        // 校验通过脉冲预清 / Verified pulse preset
_bBusyRej  := FALSE;                                                        // 忙拒预清 / Busy-rejection preset
bError     := FALSE;                                                        // 故障标志预清（R45 配对） / Error preset

(* —— 段 2：组态闸（非法即锁存） —— *)
IF _bCfgBad THEN
    _eCause := E_DL_CblCause.eCfgIllegal;                                    // 归因：组态非法 / Cause: illegal configuration
    _bFault := TRUE;                                                         // 锁存 / Latch
    _eState := E_DL_CblState.eFault;                                         // 入故障相 / Enter fault phase
END_IF

(* —— 段 3：迁出链（bReset 上升沿：清双锁存，R228B） —— *)
IF rtReset.Q THEN
    _bFault := FALSE;                                                        // 清故障锁存 / Clear fault latch
    _bFail  := FALSE;                                                        // 清标签失败锁存 / Clear the label-failure latch
    _eCause := E_DL_CblCause.eNone;                                          // 清成因 / Clear cause
    _eState := E_DL_CblState.eIdle;                                          // 回待机相 / Back to idle
END_IF

(* —— 段 4：相迁移（生成 → 打印 → 校验 握手闭环；忙时拒新） —— *)
IF (NOT _bFault) AND (NOT _bCfgBad) THEN
    CASE _eState OF

    E_DL_CblState.eIdle:
        IF rtGen.Q THEN
            IF (iLotNo < 0) OR (iLotNo > DL_CBL_LOT_MAX) THEN
                _eCause := E_DL_CblCause.eLotBad;                             // 域闸：批次号越界（信息级） / Lot out of range, info level
            ELSE
                (* 十进制拆分（每位恒 0..9，BCD 半字节合法由构造保证） *)
                _iWork := iLotNo;                                             // 取批次号 / Take the lot number
                abDigits[1] := INT_TO_BYTE(_iWork MOD 10);                    // 个位 / Units
                _iWork := _iWork / 10;                                        // 去个位 / Drop units
                abDigits[2] := INT_TO_BYTE(_iWork MOD 10);                    // 十位 / Tens
                _iWork := _iWork / 10;                                        // 去十位 / Drop tens
                abDigits[3] := INT_TO_BYTE(_iWork MOD 10);                    // 百位 / Hundreds
                _iWork := _iWork / 10;                                        // 去百位 / Drop hundreds
                abDigits[4] := INT_TO_BYTE(_iWork MOD 10);                    // 千位 / Thousands
                _uBcd := SHL(BYTE_TO_WORD(abDigits[4]), DL_CBL_SH12)
                      OR SHL(BYTE_TO_WORD(abDigits[3]), DL_CBL_SH8)
                      OR SHL(BYTE_TO_WORD(abDigits[2]), DL_CBL_SH4)
                      OR (BYTE_TO_WORD(abDigits[1]) AND DL_CBL_MSK);          // 打包 BCD / Pack BCD
                uBcdPacked := _uBcd;                                          // 打包字出口 / Packed word outlet
                _bPrintCmd := TRUE;                                           // 打印脉冲（内部位） / Internal print pulse
                _eState := E_DL_CblState.ePrinting;                           // 进打印相 / Enter printing
            END_IF
        END_IF

    E_DL_CblState.ePrinting:
        IF bPrintDone THEN
            _eState := E_DL_CblState.eVerify;                                 // 打印完成：进校验相 / Printing done, verify
        ELSIF tonPrint.Q THEN
            _bFail  := TRUE;                                                  // 打印超时：锁存 / Timeout: latch
            _bFault := TRUE;                                                  // 故障锁存 / Latch the fault
            _eCause := E_DL_CblCause.ePrintTimeout;                           // 归因：打印超时 / Cause: print timeout
            _eState := E_DL_CblState.eFault;                                  // 入故障相 / Enter fault phase
        ELSIF rtGen.Q THEN
            _bBusyRej := TRUE;                                                // 忙时拒新任务（不打断当前打印） / Busy rejection
            _eCause := E_DL_CblCause.eBusyReject;                             // 归因：忙拒（信息级） / Cause: busy rejection
        END_IF

    E_DL_CblState.eVerify:
        IF bScanValid THEN
            (* 扫码串解析：逐字符与 '0'..'9' 单字符字面量比对（ST 无字符码函数，
               故用字符串字面量判等；非法字符即判格式错） *)
            _iLen := LEN(sScanCode);                                          // 取回读长度 / Read-back length
            IF (_iLen < 1) OR (_iLen > DL_CBL_CHR_MAX) THEN
                _bFmtBad := TRUE;                                             // 长度越域：判格式错 / Length out of range
            ELSE
                _bFmtBad := FALSE;                                            // 格式结论初值 / Format result initial value
                _iVal := 0;                                                   // 数值累加器归零 / Value accumulator reset
                FOR _iPos := 1 TO DL_CBL_CHR_MAX DO
                    IF _iPos <= _iLen THEN
                        sChr := MID(sScanCode, 1, _iPos);                     // 取单个字符 / Single character
                        IF (sChr = '0') THEN
                            _iDigit := 0;
                        ELSIF (sChr = '1') THEN
                            _iDigit := 1;
                        ELSIF (sChr = '2') THEN
                            _iDigit := 2;
                        ELSIF (sChr = '3') THEN
                            _iDigit := 3;
                        ELSIF (sChr = '4') THEN
                            _iDigit := 4;
                        ELSIF (sChr = '5') THEN
                            _iDigit := 5;
                        ELSIF (sChr = '6') THEN
                            _iDigit := 6;
                        ELSIF (sChr = '7') THEN
                            _iDigit := 7;
                        ELSIF (sChr = '8') THEN
                            _iDigit := 8;
                        ELSIF (sChr = '9') THEN
                            _iDigit := 9;
                        ELSE
                            _iDigit := 0;                                     // 非法字符的数值占位（不参与累加） / Placeholder, not accumulated
                            _bFmtBad := TRUE;                                 // 非法字符 / Illegal character
                        END_IF
                        _iVal := _iVal * 10 + _iDigit;                        // 十进制累加 / Decimal accumulate
                    END_IF
                END_FOR
            END_IF

            IF _bFmtBad THEN
                _bFail  := TRUE;                                              // 格式错：锁存 / Format error: latch
                _bFault := TRUE;                                              // 故障锁存 / Latch the fault
                _eCause := E_DL_CblCause.eScanFormat;                         // 归因：回读格式非法 / Cause: scan format
                _eState := E_DL_CblState.eFault;                              // 入故障相 / Enter fault phase
            ELSIF _iVal = iLotNo THEN
                _bLabelOk := TRUE;                                            // 校验通过脉冲 / Verified pulse
                _eState := E_DL_CblState.eIdle;                               // 回待机相 / Back to idle
            ELSE
                _bFail  := TRUE;                                              // 不一致：锁存 / Mismatch: latch
                _bFault := TRUE;                                              // 故障锁存 / Latch the fault
                _eCause := E_DL_CblCause.eScanMismatch;                       // 归因：回读不一致 / Cause: scan mismatch
                _eState := E_DL_CblState.eFault;                              // 入故障相 / Enter fault phase
            END_IF
        END_IF

    E_DL_CblState.eFault:
        ;                                                                     // 故障相：仅等复位沿 / Wait for the reset edge only

    ELSE
        _eCause := E_DL_CblCause.ePhaseBad;                                   // 归因：非法相位 / Cause: illegal phase
        _bFault := TRUE;                                                      // 锁存 / Latch
        _eState := E_DL_CblState.eFault;                                      // 强拉故障相 / Force fault phase

    END_CASE
END_IF

(* —— 段 5：出口单点映射（名实双出口，R191） —— *)
bPrintCmd   := _bPrintCmd;                                                    // 打印脉冲出口 / Print pulse outlet
bLabelOk    := _bLabelOk;                                                     // 校验通过出口 / Verified outlet
bBusy       := (_eState = E_DL_CblState.ePrinting) OR (_eState = E_DL_CblState.eVerify);   // 忙碌出口 / Busy outlet
bBusyReject := _bBusyRej;                                                     // 忙拒出口 / Busy-rejection outlet
bLabelFail  := _bFail;                                                        // 标签失败出口 / Label-failure outlet
eState      := _eState;                                                       // 相出口 / Phase outlet
eCause      := _eCause;                                                       // 成因出口 / Cause outlet
bError      := _bFault;                                                       // 故障标志 / Error flag

END_FUNCTION_BLOCK
